(* IEC 61131-3 sources: STAR-PLC-Agent/results/raw/codex_matrix_resume_20261114/codex_terra/SELF008/formal/attempt_0001, 1 file *)

(* ---- candidate.st ---- *)
FUNCTION_BLOCK FB_Task
VAR_INPUT
    Request : BOOL;
    Trip : BOOL;
    Preset : USINT;
END_VAR
VAR_OUTPUT
    Ready : BOOL := FALSE;
    Count : USINT := 0;
END_VAR

IF NOT Request OR Trip OR (Preset < 1) OR (Preset > 5) THEN
    Count := 0;
    Ready := FALSE;
ELSE
    IF Count < Preset THEN
        Count := Count + 1;
    ELSE
        Count := Preset;
    END_IF;
    Ready := Count >= Preset;
END_IF;
END_FUNCTION_BLOCK
